(* IEC 61131-3 sources: Test-Git_ESME26/TestProgettoESME_26.fbsproj/PacDriveLib Migration/Motion/Homing/PDL_FB_WriteDriveEncoder.fb.st^, 5 files *)

(* ---- AsyncExtDiagTranslation.meth.st ---- *)
METHOD AsyncExtDiagTranslation : BOOL
VAR_INPUT
	i_etResult : SE_Async.ET_Result;
END_VAR

CASE i_etResult OF
	SE_Async.ET_Result.MaxNumOfReusableObjectsExceeded: ; // No error message. Try again to Start in next cycle

	SE_Async.ET_Result.AsyncAddWasNotSuccessful:
		SetDiagOutput(	i_etDiag	:= GD.ET_Diag.UnexpectedProgramBehavior,
						i_etDiagExt := PDL_ET_DiagExt.AsyncAddWasNotSuccessful,
						i_sMsg		:= SE_CTBX.FC_MultiConcat(	i_sString1 := '#',
														i_sString2 := DINT_TO_STRING(diState),
														i_sString3 := ' G_ifAsync.Start: ',
														i_sString4 := PDL_FC_EtDiagExtToString(etDiagExt)));

	SE_Async.ET_Result.InterfaceCastFailed:
		SetDiagOutput(	i_etDiag	:= GD.ET_Diag.UnexpectedProgramBehavior,
						i_etDiagExt := PDL_ET_DiagExt.InterfaceCastFailed,
						i_sMsg		:= SE_CTBX.FC_MultiConcat(	i_sString1 := '#',
														i_sString2 := DINT_TO_STRING(diState),
														i_sString3 := ' G_ifAsync.Start: ',
														i_sString4 := PDL_FC_EtDiagExtToString(etDiagExt)));

	SE_Async.ET_Result.SemaphoreCreateFailed:
		SetDiagOutput(	i_etDiag	:= GD.ET_Diag.UnexpectedProgramBehavior,
						i_etDiagExt := PDL_ET_DiagExt.SemaphoreMeCreateFailed,
						i_sMsg		:= SE_CTBX.FC_MultiConcat(	i_sString1 := '#',
														i_sString2 := DINT_TO_STRING(diState),
														i_sString3 := ' G_ifAsync.Start: ',
														i_sString4 := PDL_FC_EtDiagExtToString(etDiagExt)));

	SE_Async.ET_Result.AsyncInvalid:
		SetDiagOutput(	i_etDiag	:= GD.ET_Diag.InputParameterInvalid,
						i_etDiagExt := PDL_ET_DiagExt.AsyncInvalid,
						i_sMsg		:= SE_CTBX.FC_MultiConcat(	i_sString1 := '#',
														i_sString2 := DINT_TO_STRING(diState),
														i_sString3 := ' G_ifAsync.Start: ',
														i_sString4 := PDL_FC_EtDiagExtToString(etDiagExt)));

	SE_Async.ET_Result.NoAsyncTasksCreated:
		SetDiagOutput(	i_etDiag	:= GD.ET_Diag.ExecutionAborted,
						i_etDiagExt := PDL_ET_DiagExt.NoAsyncTasksCreated,
						i_sMsg		:= SE_CTBX.FC_MultiConcat(	i_sString1 := '#',
														i_sString2 := DINT_TO_STRING(diState),
														i_sString3 := ' G_ifAsync.Start: ',
														i_sString4 := PDL_FC_EtDiagExtToString(etDiagExt)));

	SE_Async.ET_Result.AsyncInitNotFinished:
		SetDiagOutput(	i_etDiag	:= GD.ET_Diag.ExecutionAborted,
						i_etDiagExt := PDL_ET_DiagExt.AsyncInitNotFinished,
						i_sMsg		:= SE_CTBX.FC_MultiConcat(	i_sString1 := '#',
														i_sString2 := DINT_TO_STRING(diState),
														i_sString3 := ' G_ifAsync.Start: ',
														i_sString4 := PDL_FC_EtDiagExtToString(etDiagExt)));

	SE_Async.ET_Result.ColdResetOfControllerNecessary:
		SetDiagOutput(	i_etDiag	:= GD.ET_Diag.ExecutionAborted,
						i_etDiagExt := PDL_ET_DiagExt.ColdResetOfControllerNecessary,
						i_sMsg		:= SE_CTBX.FC_MultiConcat(	i_sString1 := '#',
														i_sString2 := DINT_TO_STRING(diState),
														i_sString3 := ' G_ifAsync.Start: ',
														i_sString4 := PDL_FC_EtDiagExtToString(etDiagExt)));

	ELSE
		SetDiagOutput(	i_etDiag	:= GD.ET_Diag.UnexpectedProgramBehavior,
						i_etDiagExt := PDL_ET_DiagExt.UnexpectedFeedback,
						i_sMsg		:= SE_CTBX.FC_MultiConcat(	i_sString1 := '#',
														i_sString2 := DINT_TO_STRING(diState),
														i_sString3 := ' G_ifAsync.Start: ',
														i_sString4 := PDL_FC_EtDiagExtToString(etDiagExt)));
END_CASE

(* ---- AverageVel.meth.st ---- *)
{attribute 'hide'}
METHOD AverageVel : BOOL
VAR_INPUT
END_VAR
VAR
END_VAR

AverageVel := TRUE;

lrSum		:= lrSum + i_ifDrive.RefVelocity - alrA[uiI];	(* lrSum = lrSum + New Value - Oldest Value *)
alrA[uiI]	:= i_ifDrive.RefVelocity ;
uiI			:= uiI + 1;
lrAverage	:= lrSum / 16;

IF uiI > 16 THEN
	uiI		:= 1;
	xValid	:= TRUE;
END_IF

(* ---- ParameterCheckEnable.meth.st ---- *)
METHOD PRIVATE ParameterCheckEnable : BOOL

VAR
	ifGetParentDevice      : DTSI.IF_GetParentDevice;
	ifDeviceAccess         : DTSI.IF_DeviceAccess;
END_VAR

diSercosState := FC_GetSercosState();

IF diSercosState <> 4 THEN
	SetDiagOutput(	i_etDiag	:= GD.ET_Diag.SercosConditionInvalid,
					i_etDiagExt := PDL_ET_DiagExt.SercosNotInPhaseFour,
					i_sMsg		:= '');
	RETURN;
END_IF

IF i_ifDrive = 0 THEN
	SetDiagOutput(	i_etDiag	:= GD.ET_Diag.InputParameterInvalid,
					i_etDiagExt := PDL_ET_DiagExt.DriveInvalid,
					i_sMsg		:= 'i_ifDrive - Invalid Interface');
	RETURN;
END_IF

xSuccess := __QUERYINTERFACE(i_ifDrive, ifGetParentDevice);
IF NOT xSuccess OR ifGetParentDevice = 0 THEN
	SetDiagOutput(	i_etDiag	:= GD.ET_Diag.InputParameterInvalid,
					i_etDiagExt := PDL_ET_DiagExt.DriveInvalid,
					i_sMsg		:= 'i_ifDrive - IF_GetParentDevice not implemented.');
	RETURN;
END_IF

ifDeviceAccess := ifGetParentDevice.GetParentDevice();

xSuccess := __QUERYINTERFACE(ifDeviceAccess,ifScalingAccess );
IF (NOT xSuccess OR ifScalingAccess = 0) THEN
	SetDiagOutput(	i_etDiag	:= GD.ET_Diag.InputParameterInvalid,
					i_etDiagExt := PDL_ET_DiagExt.DriveInvalid,
					i_sMsg		:= 'i_ifDrive - IF_Scaling not implemented.');
	RETURN;
END_IF
ifScaling := ifScalingAccess.Scaling;

xSuccess := __QUERYINTERFACE(ifDeviceAccess,ifDriveAccess );
IF (NOT xSuccess OR ifDriveAccess = 0) THEN
	q_etDiag	:= GD.ET_Diag.InputParameterInvalid;
	q_etDiagExt := PDL_ET_DiagExt.DriveInvalid;
	q_sMsg		:= 'i_ifDrive - IF_Drive not implemented.';
	RETURN;
END_IF
ifDrive := ifDriveAccess.Drive;

xSuccess := __QUERYINTERFACE(ifDeviceAccess,ifDrive2Access );
IF (NOT xSuccess OR ifDrive2Access = 0) THEN
	q_etDiag	:= GD.ET_Diag.InputParameterInvalid;
	q_etDiagExt := PDL_ET_DiagExt.DriveInvalid;
	q_sMsg		:= 'i_ifDrive - IF_Drive2 not implemented.';
	RETURN;
END_IF
ifDrive2 := ifDrive2Access.Drive2;

xSuccess := __QUERYINTERFACE(ifDeviceAccess,ifDriveConfigAccess );
IF (NOT xSuccess OR ifDriveConfigAccess = 0) THEN
	q_etDiag	:= GD.ET_Diag.InputParameterInvalid;
	q_etDiagExt := PDL_ET_DiagExt.DriveInvalid;
	q_sMsg		:= 'i_ifDrive - IF_Drive not implemented.';
	RETURN;
END_IF
ifDriveConfig := ifDriveConfigAccess.DriveConfig;

xSuccess := __QUERYINTERFACE(ifDeviceAccess,ifMotorAccess );
IF (NOT xSuccess OR ifMotorAccess = 0) THEN
	SetDiagOutput(	i_etDiag	:= GD.ET_Diag.InputParameterInvalid,
					i_etDiagExt := PDL_ET_DiagExt.DriveInvalid,
					i_sMsg		:= 'i_ifDrive - IF_Motor not implemented.');
	diState := 0;
	RETURN;
END_IF
ifMotor := ifMotorAccess.Motor;

xSuccess := __QUERYINTERFACE(ifDeviceAccess,ifEncoderAccess );
IF (NOT xSuccess OR ifEncoderAccess = 0) THEN
	SetDiagOutput(	i_etDiag	:= GD.ET_Diag.InputParameterInvalid,
					i_etDiagExt := PDL_ET_DiagExt.DriveInvalid,
					i_sMsg		:= 'i_ifDrive - IF_Encoder not implemented.');
	diState := 0;
	RETURN;
END_IF
ifEncoder := ifEncoderAccess.Encoder;

xSuccess := __QUERYINTERFACE(ifDeviceAccess,ifLXM62DriveAccess );
IF (NOT xSuccess OR ifLXM62DriveAccess = 0) THEN
	SetDiagOutput(	i_etDiag	:= GD.ET_Diag.InputParameterInvalid,
					i_etDiagExt := PDL_ET_DiagExt.DriveInvalid,
					i_sMsg		:= 'i_ifDrive - IF_LXM62DriveAccess not implemented.');
	diState := 0;
	RETURN;
END_IF
ifLXM62Drive := ifLXM62DriveAccess.Lexium62Drive;

xSuccess := __QUERYINTERFACE(ifDeviceAccess, ifWorkingModeAccess);
IF (NOT xSuccess OR ifLXM62DriveAccess = 0) THEN
	SetDiagOutput(	i_etDiag	:= GD.ET_Diag.InputParameterInvalid,
					i_etDiagExt := PDL_ET_DiagExt.DriveInvalid,
					i_sMsg		:= 'i_ifDrive - IF_LXM62DriveAccess not implemented.');
	RETURN;
END_IF
ifWorkingMode := ifWorkingModeAccess.WorkingMode;

xSuccess := __QUERYINTERFACE(ifDeviceAccess, ifDeviceType);
IF (NOT xSuccess OR ifDeviceType = 0) THEN
	SetDiagOutput(	i_etDiag	:= GD.ET_Diag.InputParameterInvalid,
					i_etDiagExt := PDL_ET_DiagExt.DriveInvalid,
					i_sMsg 		:= 'i_ifDrive - IF_Device_Type not implemented');
	diState := 0;
	RETURN;
END_IF

lrEncoderRange := ifEncoder.Revolutions;
IF (ABS(lrEncoderRange) < 1.0E-3) THEN
	SetDiagOutput(	i_etDiag	:= GD.ET_Diag.DriveConditionInvalid,
					i_etDiagExt := PDL_ET_DiagExt.DriveEncoderInvalid,
					i_sMsg		:= '');
	RETURN;
ELSE
	lrEncoderPeriode := ifEncoder.Revolutions * ifScaling.PositionResolution * TO_LREAL(ifScaling.GearIn) / TO_LREAL(ifScaling.GearOut);
END_IF

IF (ifWorkingMode.ActualState <> CFDI.ET_WorkingState.Physical) THEN		// prüfen, ob Achse real und Motor angeschlossen
	SetDiagOutput(	i_etDiag	:= GD.ET_Diag.DriveConditionInvalid,
					i_etDiagExt := PDL_ET_DiagExt.NoRealDrive,
					i_sMsg		:= '');
	RETURN;
ELSIF (i_lrUserPeriod < 0.0) THEN
	SetDiagOutput(	i_etDiag	:= GD.ET_Diag.InputParameterInvalid,
					i_etDiagExt := PDL_ET_DiagExt.UserPeriodRange,
					i_sMsg		:= '0.0 <= i_lrUserPeriod');
	RETURN;
ELSIF (i_lrUserPeriod < c_lrRealNull) AND ( (i_lrAbsEncOffset < c_lrRealNull) OR (i_lrAbsEncOffset > (lrEncoderPeriode - c_lrRealNull)) ) THEN
	SetDiagOutput(	i_etDiag	:= GD.ET_Diag.InputParameterInvalid,
					i_etDiagExt := PDL_ET_DiagExt.AbsEncOffsetRange,
					i_sMsg		:= STANDARD.CONCAT('0.0 < i_lrAbsEncOffset <= ', SE_CTBX.FC_LrealToString(i_sFormat := '#0.00', i_lrInput := lrEncoderPeriode - c_lrRealNull) ));
	RETURN;
(* Check if UserPeriode fits into EncoderPeriode *)
ELSIF(i_lrUserPeriod > c_lrRealNull) AND ( ABS(lrEncoderPeriode/i_lrUserPeriod - TRUNC_INT(lrEncoderPeriode / i_lrUserPeriod)) > c_lrRealNull ) THEN
	SetDiagOutput(	i_etDiag	:= GD.ET_Diag.InputParameterInvalid,
					i_etDiagExt := PDL_ET_DiagExt.UserPeriodRange,
					i_sMsg		:= STANDARD.CONCAT('i_lrUserPeriod has to be a divsior of ', SE_CTBX.FC_LrealToString(i_sFormat := '#0.00', i_lrInput := lrEncoderPeriode)));
	RETURN;
END_IF

ParameterCheckEnable := TRUE;

(* ---- SetDiagOutput.meth.st ---- *)
{attribute 'hide'}
METHOD SetDiagOutput : BOOL
VAR_INPUT
	i_etDiag	: GD.ET_Diag;
	i_etDiagExt	: PDL_ET_DiagExt;
	i_sMsg		: STRING[80];
END_VAR
VAR
END_VAR

IF q_etDiag = GD.ET_Diag.OK OR i_etDiagExt = PDL_ET_DiagExt.Disabled THEN

	q_etDiag 	:= i_etDiag;
	q_etDiagExt := i_etDiagExt;
	q_sMsg 		:= i_sMsg;

END_IF

(* ---- WritePosition.meth.st ---- *)
METHOD INTERNAL WritePosition

CASE diWritePositionState OF

10:
	IF i_lrUserPeriod > c_lrRealNull THEN
		lrModuloPosition := lrEncoderPeriode / 2.0 + i_ifDrive.RefPosition - lrSavePosition;
	ELSE
		lrModuloPosition := i_lrAbsEncOffset + i_ifDrive.RefPosition - lrSavePosition;
	END_IF

	IF ifScaling.InvertDirection = FALSE THEN // Motor direction right
		lrPositionTemp	:= lrModuloPosition;
	ELSE
		lrPositionTemp := lrEncoderPeriode - lrModuloPosition;
	END_IF

	// Execute after increasing cycle-time or asynchronous
	fbSetDrvEncPos.ifDeviceType					:= ifDeviceType;
	fbSetDrvEncPos.lrPosition				:= lrPositionTemp;

	SE_Async.G_ifAsyncMgr.Start(
		i_ifAsync    := fbSetDrvEncPos,
		q_etResult   => etResult,
		q_sResultMsg => sResultMsg,
		q_xError     => xError);

	IF xError THEN
		AsyncExtDiagTranslation(i_etResult := etResult);
		RETURN;
	ELSE
		diWritePositionState := 20;
	END_IF

20:
	IF fbSetDrvEncPos.xDone THEN
		diWritePositionState := 30;
	END_IF

30:	// Check Result of writing
	diResult := fbSetDrvEncPos.diResultSetDrvEncPos;
	IF diResult = 0  THEN // Ok
		tonTimeOut(IN := FALSE, PT := c_timProgramTime );

		SetDiagOutput(	i_etDiag	:= GD.ET_Diag.Ok,
						i_etDiagExt := PDL_ET_DiagExt.WaitUntilEncoderWritten,
						i_sMsg		:= '');
		diState	:= 20;
	ELSIF diResult = -3 THEN
		SetDiagOutput(	i_etDiag	:= GD.ET_Diag.InputParameterInvalid,
						i_etDiagExt := PDL_ET_DiagExt.DriveInvalid,
						i_sMsg		:= 'Drive must not be virtual');
		diState := 0;
	ELSIF diResult = -4 THEN
		SetDiagOutput(	i_etDiag	:= GD.ET_Diag.InputParameterInvalid,
						i_etDiagExt := PDL_ET_DiagExt.DriveInvalid,
						i_sMsg		:= 'Drive must not be deactivated');
		diState := 0;
	ELSE	(* Programming error *)
		SetDiagOutput(	i_etDiag	:= GD.ET_Diag.UnexpectedProgramBehavior,
						i_etDiagExt := PDL_ET_DiagExt.UnexpectedFeedback,
						i_sMsg		:= CONCAT('FC_DrvEncSetPosition: ', DINT_TO_STRING(diResult)));
		q_xReady := FALSE;
		diState	:= 0;
	END_IF

END_CASE
